Fanuc KAREL source: KA00005.KL

PROGRAM KA00005
%NOLOCKGROUP
VAR
  SRC: INTEGER
  DST: POSITION
BEGIN
  SRC = 2
  DST = SRC
END KA00005
